(*
SPDX-FileCopyrightText: © 2026 Oleksandr Tiutyk <trofimich@gmail.com>
SPDX-License-Identifier: MIT
License: https://opensource.org/license/mit
*)

(*!
<summary>Holds a single-field structure for explicit VAR_INFO type resolution.</summary>
*)
TYPE JSON_TEST_SINGLE_VALUE :
STRUCT
	//! <summary>Value restored through the explicit structure type.</summary>
	Number : DINT;
END_STRUCT
END_TYPE

(* stored: Version 1.1.0.1
   DUT JSON_TEST_SINGLE_VALUE: Id {6e657c52-7e31-4780-9099-cd46aa4156a7} *)
